Fanuc KAREL source: kt00409.KL

-- PROVISIONAL review KL for V770-1; original PC SHA256 5d74139c3ed6186f3529df50e07a04ea052c324933dbd4ac5d7ea49cdc43371a
-- Incomplete behavior may be omitted. Consult companion uncertainty JSON. Do not deploy.
PROGRAM KT00409
%NOLOCKGROUP
VAR
  B1 : BOOLEAN
  B2 : BOOLEAN
  OUT : BOOLEAN
BEGIN
  -- UNRESOLVED_PC offsets 5-12; opcodes 9D,23
  -- UNRESOLVED_PC offsets 17-24; opcodes 9C,23
  -- UNRESOLVED_PC offsets 29-36; opcodes 9D,23
  -- UNRESOLVED_PC offsets 41-48; opcodes 9C,23
  -- UNRESOLVED_PC offsets 53-72; opcodes 21,21,5B,23
  -- UNRESOLVED_PC offsets 77-81; opcodes 7F
END KT00409
